Fanuc KAREL source: ko00057.KL

-- PROVISIONAL review KL for V1013-1; original PC SHA256 4b2e1ae0924b5d394569b1ab30afa0e8c33bb1069f99e6895a1b308231c0a856
-- Incomplete behavior may be omitted. Consult companion uncertainty JSON. Do not deploy.
PROGRAM KO00057
%NOLOCKGROUP
BEGIN
  -- UNRESOLVED_PC offsets 5-12; opcodes 9D,23
  -- UNRESOLVED_PC offsets 17-69; opcodes 27,27,49,7E,AD,27,49,7E,AD,22,31,7E,4A
  -- UNRESOLVED_PC offsets 74-78; opcodes 7F
END KO00057
